// TIA Portal V20 export
DATA_BLOCK "T6_Resultado"   // DB43901
{ S7_Optimized_Access := 'TRUE' }
AUTHOR : IA
FAMILY : PRUEBA
VERSION : 0.1
// Tanda 2: un Bool por prueba
// stored: AutoNumber false
   VAR
      L_T_CONV_T_DI : Bool;   // T_CONV Time→DInt
      L_T_CONV_DI_T : Bool;   // T_CONV DInt→Time
      L_T_ADD : Bool;   // T_ADD DTL + Time (10:00 + 1h)
      L_T_SUB : Bool;   // T_SUB DTL − Time (10:00 − 1h)
      L_T_DIFF : Bool;   // T_DIFF DTL (11:00 − 10:00)
      L_T_COMBINE : Bool;   // T_COMBINE Date + Time_Of_Day
      L_RD_LOC_T : Bool;   // RD_LOC_T (hora local)
      L_WR_LOC_T : Bool;   // WR_LOC_T
      L_WR_SYS_T : Bool;   // WR_SYS_T
      L_Eq_DTL : Bool;   // Eq con SrcType DTL
      L_S_CONV_I_S : Bool;   // S_CONV Int→String (comprobado con la vuelta)
      L_S_CONV_S_I : Bool;   // S_CONV String→Int
      L_LEFT : Bool;   // LEFT
      L_RIGHT : Bool;   // RIGHT
      L_MID : Bool;   // MID
      L_DELETE : Bool;   // DELETE
      L_INSERT : Bool;   // INSERT
      L_REPLACE : Bool;   // REPLACE
      L_FIND : Bool;   // FIND
      L_ATH : Bool;   // ATH '1A2B' → 16#1A, 16#2B
      L_HTA : Bool;   // HTA 16#1A, 16#2B → '1A2B'
      L_Eq_Char : Bool;   // Eq con SrcType Char
      S_Fecha : Bool;   // [SCL] TIME_TO_DINT, DINT_TO_TIME, T_ADD, T_SUB, T_DIFF, CONCAT_DATE_TOD (T_COMBINE en KOP)
      S_Reloj : Bool;   // [SCL] RD_LOC_T, RD_SYS_T, WR_LOC_T y WR_SYS_T (una vez)
      S_Texto : Bool;   // [SCL] INT_TO_STRING, STRING_TO_INT, LEFT, RIGHT, MID, DELETE, INSERT, REPLACE, FIND
      S_Hex : Bool;   // [SCL] ATH y HTA
      S_Comparar : Bool;   // [SCL] comparar DTL y Char
      Vida : DInt;   // Sube cada ciclo
      OK : Int;   // Correctas
      Total : Int := 27;   // Pruebas
      Todo_OK : Bool;   // Todas correctas
   END_VAR
BEGIN
END_DATA_BLOCK
